(* IEC 61131-3 sources: Elmo_Master/Lasal_PRG/Elmo_EtherCAT_Test_4Axis/Class/EtherCAT_SDOBase, 1 file *)

(* ---- EtherCAT_SDOBase.st ---- *)
#include "..\..\Class\ECAT_Master_Base\ECAT_Master_Base.h"

(*!
<Class
	Name               = "EtherCAT_SDOBase"
	Revision           = "1.1"
	RealtimeTask       = "false"
	CyclicTask         = "false"
	BackgroundTask     = "false"
	Sigmatek           = "true"
	OSInterface        = "false"
	HighPriority       = "false"
	Automatic          = "false"
	UpdateMode         = "Prescan"
	IconPath           = ".\Class\EtherCAT.ico"
	SharedCommandTable = "true"
	Objectsize         = "(510,120)"
	Comment            = "Class can be used to establish a SDO Communication with an EtherCAT slave module.">
	<Channels>
		<Server Name="ClassState" Visualized="true" Initialize="false" WriteProtected="true" Retentive="false" Comment="Shows the state of the class."/>
		<Server Name="CompleteAccess" Visualized="true" Initialize="true" DefValue="0" WriteProtected="false" Retentive="false" Comment="Accesstype of the SDO.&#13;&#10;0 .. Single Access&#13;&#10;1 .. Complete Access"/>
		<Server Name="ErrorCode" Visualized="true" Initialize="false" WriteProtected="true" Retentive="false" Comment="Shows the Errorcode of the SDO handling if ClassState = ERROR.&#13;&#10;&#13;&#10;0x05030000 ... toggle bit not changed&#13;&#10;0x05040000 ...  SDO protocol timeout&#13;&#10;0x05040001 ...  SDO command specifier invalid or unknown&#13;&#10;0x05040005 ...  not enough space in the main memory&#13;&#10;0x06010000 ...  access to this object is not supported&#13;&#10;0x06010001 ...  attempt to read to a write_only parameter&#13;&#10;0x06010002 ...  attempt to write to a read_only parameter&#13;&#10;0x06010003 ...  SubIdx 0 can only be written if it is 0&#13;&#10;0x06010004 ...  SDO complete access is not supported for ENUMs&#13;&#10;0x06010005 ...  object length is larger than mailbox size&#13;&#10;0x06010006 ...  object mapped to RxPDO, SDO download blocked&#13;&#10;0x06020000 ...  the object is not found in the object directory&#13;&#10;0x06040041 ...  object can&apos;t be mapped in the PDO&#13;&#10;0x06040042 ...  the amount and length of objects exceeds the PDO length&#13;&#10;0x06040043 ...  general parameter incompatibility reason&#13;&#10;0x06040047 ...  general internal incompatibility in the device&#13;&#10;0x06060000 ...  access failed due to a hardware error&#13;&#10;0x06070000 ...  data type does not match, length of service parameter does not match&#13;&#10;0x06070012 ...  data type does not match, length of service parameter too high&#13;&#10;0x06070013 ...  data type does not match, length of service parameter too low&#13;&#10;0x06090011 ...  sub index does not exist&#13;&#10;0x06090030 ...  value of range of parameter exceeded (only for write access)&#13;&#10;0x06090031 ...  value of range of parameter too high&#13;&#10;0x06090032 ...  value of range of parameter to low&#13;&#10;0x06090036 ...  maximum value is less than minimum value&#13;&#10;0x08000000 ...  general error&#13;&#10;0x08000020 ...  data can&apos;t be stored to the application&#13;&#10;0x08000021 ...  data can&apos;t be stored to the application because of local control&#13;&#10;0x08000022 ...  data can&apos;t be stored to the application because of present device state&#13;&#10;0x08000023 ...  object dictionary dynamic generation failed or no object dict. is present"/>
		<Server Name="ParaIndex" Visualized="true" Initialize="true" WriteProtected="false" Retentive="false" Comment="Index from the SDO Entry"/>
		<Server Name="ParaLength" Visualized="true" Initialize="true" WriteProtected="false" Retentive="false" Comment="ParaReadWrite = 0&#13;&#10;Shows the amount of data bytes which were read.&#13;&#10;&#13;&#10;ParaReadWrite = 1&#13;&#10;The set amount of data bytes will be written to the parameter. (not necessary if ParaType = 1)"/>
		<Server Name="ParaReadWrite" Visualized="true" Initialize="true" WriteProtected="false" Retentive="false" Comment="Read or Write the set parameter.&#13;&#10;0 .. Read&#13;&#10;1 .. Write"/>
		<Server Name="ParaString" Class="String" Visualized="true" Initialize="true" WriteProtected="false" Retentive="false" Comment="Shows the value of the parameter as a String (if ParaType = 1)."/>
		<Server Name="ParaSubIndex" Visualized="true" Initialize="true" WriteProtected="false" Retentive="false" Comment="Subindex from the SDO Entry"/>
		<Server Name="ParaType" Visualized="true" Initialize="true" WriteProtected="false" Retentive="false" Comment="The type of the parameter can be set with this server&#13;&#10;0 ... Value&#13;&#10;1 ... String"/>
		<Server Name="ParaValue" Visualized="true" Initialize="true" WriteProtected="false" Retentive="false" Comment="Value of the set parameter.&#13;&#10;&#13;&#10;ParaReadWrite = 0&#13;&#10;Shows the value of the read parameter.&#13;&#10;&#13;&#10;ParaReadWrite = 1&#13;&#10;The value of this server will be written to the set parameter."/>
		<Server Name="Timeout" Visualized="true" Initialize="true" DefValue="100" WriteProtected="false" Retentive="false" Comment="Maximum time before SDO handling generates an error in ms. (Default = 100)"/>
		<Client Name="strSDOParaString" Required="true" Internal="true"/>
		<Client Name="toSlave" Required="true" Internal="false" Comment="Has to be connected to the ClassState server of an Ethercat slave module."/>
	</Channels>
	<Dependencies>
		<Files>
			<File Path=".\Class\ECAT_Master_Base\ECAT_Master_Base.h" Include="true"/>
		</Files>
	</Dependencies>
	<RevDoku>
		<Owner Company="Sigmatek" Author="EisMic"/>
		<Dokumentation Revision="1.1" Date="2026-02-20" Author="WinPat" Company="Sigmatek" Description="Replaced the GetDataAt() Method with the TxtGet() Method, when Reading a String, to prevent faulty results, when the new String is shorter than the string that was written before"/>
		<Dokumentation Revision="1.0" Date="09.04.2020" Author="EisMic" Company="Sigmatek" Description="First release version."/>
		<Dokumentation Revision="0.1" Date="17.05.2019" Author="EisMic" Company="Sigmatek" Description="First test version."/>
	</RevDoku>
	<Network Name="EtherCAT_SDOBase">
		<!-- List of Components in this network -->
		<Components>
			<Object
				Name       = "strSDOParaString"
				Class      = "String"
				Position   = "(150,600)"
				Visualized = "true"
				Remotely   = "true">
				<Channels>
					<Server Name="Data"/>
					<Client Name="SingleRealloc" Value="1"/>
				</Channels>
			</Object>
		</Components>
		<Comments>
		</Comments>
		<!-- List of Connections in this network -->
		<Connections>
			<Connection Source="this.strSDOParaString" Destination="strSDOParaString.Data"/>
			<Connection Source="this.ParaString" Destination="strSDOParaString.Data" Vertices="(638,690),(466,690),"/>
		</Connections>
		<!-- Headerfiles -->
		<Options>
		</Options>
	</Network>
</Class>
*)
EtherCAT_SDOBase : CLASS
  //Servers:
	ClassState 	: SvrChCmd_iprStates;
	ParaReadWrite 	: SvrCh_DINT;
	ParaIndex 	: SvrCh_HDINT;
	ParaSubIndex 	: SvrCh_HDINT;
	CompleteAccess 	: SvrCh_DINT;
	ParaType 	: SvrCh_DINT;
	ParaLength 	: SvrCh_UDINT;
	ParaValue 	: SvrCh_DINT;
	ParaString 	: SvrChCmd_UDINT;
	ErrorCode 	: SvrCh_HDINT;
	Timeout 	: SvrCh_UDINT;
  //Clients:
	toSlave 	: CltChCmd_ECAT_Slave_Base;
	strSDOParaString 	: CltChCmd_String;
  //Variables:
		szString : ARRAY [0..199] OF CHAR;

  //Functions:

	FUNCTION VIRTUAL GLOBAL ClassState::NewInst
		VAR_INPUT
			pPara 	: ^CmdStruct;
			pResult 	: ^results;
		END_VAR
		VAR_OUTPUT
			ret_code 	: iprStates;
		END_VAR;

	FUNCTION VIRTUAL GLOBAL ParaReadWrite::Write
		VAR_INPUT
			input (EAX) 	: DINT;
		END_VAR
		VAR_OUTPUT
			result (EAX) 	: DINT;
		END_VAR;

	FUNCTION VIRTUAL GLOBAL ParaType::Write
		VAR_INPUT
			input (EAX) 	: DINT;
		END_VAR
		VAR_OUTPUT
			result (EAX) 	: DINT;
		END_VAR;

	FUNCTION VIRTUAL GLOBAL ParaString::Read
		VAR_OUTPUT
			output (EAX) 	: UDINT;
		END_VAR;

	FUNCTION VIRTUAL GLOBAL ParaString::Write
		VAR_INPUT
			input (EAX) 	: UDINT;
		END_VAR
		VAR_OUTPUT
			result (EAX) 	: UDINT;
		END_VAR;
  //Tables:
	FUNCTION @STD
		VAR_OUTPUT
			ret_code	: CONFSTATES;
		END_VAR;
	FUNCTION GLOBAL TAB @CT_;
END_CLASS;

#pragma using String
#pragma usingLtd ECAT_Slave_Base

FUNCTION VIRTUAL GLOBAL EtherCAT_SDOBase::ParaReadWrite::Write
	VAR_INPUT
		input (EAX) 	: DINT;
	END_VAR
	VAR_OUTPUT
		result (EAX) 	: DINT;
	END_VAR
  VAR
  	retcode : iprStates;
  END_VAR

	ParaReadWrite := input;
	result := ParaReadWrite;

  // check if the class is ready is ready for a new asy command
  if (ClassState <> BUSY) then

    //Check for Read or Write Para
    if ParaReadWrite = 0 then

      //Read Parameter

      //Check if value or string (0 .. value, 1 .. string)
      if ParaType = 0 then
        ParaValue := 0;
        retcode := toSlave.StartReadSDO(ParaIndex$HINT,ParaSubIndex$HSINT,CompleteAccess,(#ParaValue)$^USINT,sizeof(ParaValue),Timeout,THIS);
      else
        strSDOParaString.Clear();
        retcode := toSlave.StartReadSDO(ParaIndex$HINT,ParaSubIndex$HSINT,CompleteAccess,(#szString)$^USINT,SIZEOF(szString),Timeout,THIS);
      end_if;
    else

      //Write parameter

      //Check if value or string (0 .. value, 1 .. string)
      if ParaType = 0 then
        retcode := toSlave.StartWriteSDO(ParaIndex$HINT,ParaSubIndex$HSINT,CompleteAccess,(#ParaValue)$^USINT,ParaLength,Timeout,THIS);
      else
        ParaLength := strSDOParaString.GetLength() + strSDOParaString.GetCharSize();
        strSDOParaString.TxtGet(pdst:=#szString[0], dstsize:=sizeof(szString));
        retcode := toSlave.StartWriteSDO(ParaIndex$HINT,ParaSubIndex$HSINT,CompleteAccess,#szString[0],ParaLength,Timeout,THIS);
      end_if;
    end_if;

    if retcode = READY then
      ClassState := BUSY; //Show that SDO is busy
    else
      ClassState := ERROR;
    end_if;
  end_if;

END_FUNCTION

FUNCTION VIRTUAL GLOBAL EtherCAT_SDOBase::ParaString::Read
	VAR_OUTPUT
		output (EAX) 	: UDINT;
	END_VAR

	ParaString := strSDOParaString.Data.Read();
	output := ParaString;

END_FUNCTION

FUNCTION VIRTUAL GLOBAL EtherCAT_SDOBase::ParaString::Write
	VAR_INPUT
		input (EAX) 	: UDINT;
	END_VAR
	VAR_OUTPUT
		result (EAX) 	: UDINT;
	END_VAR

	ParaString := input;
	result := (strSDOParaString.Data.Write(ParaString))$UDINT;

END_FUNCTION

FUNCTION VIRTUAL GLOBAL EtherCAT_SDOBase::ClassState::NewInst
	VAR_INPUT
		pPara 	: ^CmdStruct;
		pResult 	: ^Results;
	END_VAR
	VAR_OUTPUT
		ret_code 	: IprStates;
	END_VAR

	CASE pPara^.uiCmd OF
// *******************************************************************************
		ECAT_M_SDO_CALLBACK: // succeeded to get/set value

      if pPara^.aPara[0]$DINT = 1 then //Check version

        //Check return code
        if pPara^.aPara[1]$DINT = 0 then

          //Read SDO
          if pPara^.aPara[2]$BOOL = 0 then

            ParaLength := pPara^.aPara[5]$UDINT;

            //Write string to string object (if Paratype = 0 Value is already written to server)
            if ParaType = 1 then
              strSDOParaString.TxtSet(dstchrsize:=1, psrc:=#szString[0], srcchrsize:=1);
            end_if;

            ClassState := READY;
            ErrorCode  := 0;

          //Write SDO
          elsif pPara^.aPara[2]$BOOL = 1 then

            //Write para was succesfull
            ClassState := READY;
            ErrorCode  := 0;

          else
            //Invalid command
            ClassState := ERROR;
          end_if;
       else
          ErrorCode := pPara^.aPara[6]$UDINT;
          //Error
          ClassState := ERROR;
        end_if;
      else
        //Invalid version
        ClassState := ERROR;
      end_if;

	END_CASE;

	ret_code := READY;

END_FUNCTION

FUNCTION VIRTUAL GLOBAL EtherCAT_SDOBase::ParaType::Write
	VAR_INPUT
		input (EAX) 	: DINT;
	END_VAR
	VAR_OUTPUT
		result (EAX) 	: DINT;
	END_VAR

  if input = 0 then
    ParaType := 0;
  else
    ParaType := 1;
  end_if;

	result := ParaType;

END_FUNCTION
